Universal Robots URScript: FeedConveyor.script

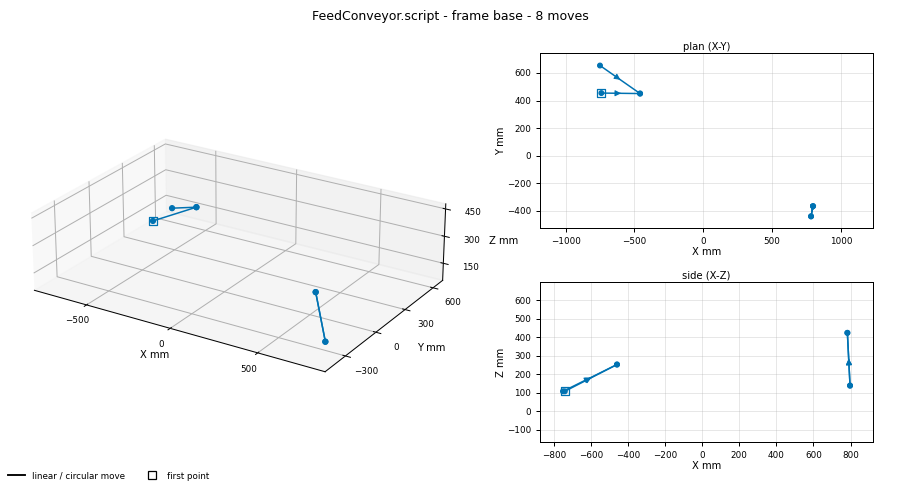
[picture p0: tool path of FeedConveyor.script in frame base, 8 of 12 moves have a stored position in this frame; points joined in program order, loops and branches not executed]
def FeedConveyor():
  # Global parameters:
  global speed_ms    = 0.250
  global speed_rads  = 0.750
  global accel_mss   = 1.200
  global accel_radss = 1.200
  global blend_radius_m = 0.001
  global ref_frame = p[0,0,0,0,0,0]

  #
  # TO REMOVE HEADER:
  # Go to "Program" -> "Post-Processor Editor"
  # Select "Universal Robots"
  # Set "INCLUDE_HEADER" to "False"
  #
  #--------------------------
  # Add any default subprograms here
  # For example, to drive a gripper as a program call:
  # def Gripper_Open():
  #   ...
  # end
  #
  # Example to drive a spray gun:
  def SprayOn(value):
    # use the value as an output:
    DO_SPRAY = 5
    if value == 0:
      set_standard_digital_out(DO_SPRAY, False)
    else:
      set_standard_digital_out(DO_SPRAY, True)
    end
  end

  # Example to drive an extruder:
  def Extruder(value):
    # use the value as an output:
    if value < 0:
      # stop extruder
    else:
      # start extruder
    end
  end

  # Example to move an external axis
  def MoveAxis(value):
    # use the value as an output:
    DO_AXIS_1 = 1
    DI_AXIS_1 = 1
    if value <= 0:
      set_standard_digital_out(DO_AXIS_1, False)

      # Wait for digital input to change state
      #while (get_standard_digital_in(DI_AXIS_1) != False):
      #  sync()
      #end
    else:
      set_standard_digital_out(DO_AXIS_1, True)

      # Wait for digital input to change state
      #while (get_standard_digital_in(DI_AXIS_1) != True):
      #  sync()
      #end
    end
  end
  #--------------------------


  # Main program:
  # Program generated by VerticalBot Studio for UR10 A on 25/10/2026 12:00:00
  # Using nominal kinematics.
  ref_frame = p[-1.052120, 0.561703, 0.068352, 0.000000, 0.000000, 1.570796]
  set_tcp(p[0.000000, -0.020000, 0.130000, 0.000000, 0.000000, 0.000000])
  movej([-1.414502, -1.531893, 2.172743, -0.640850, 0.156295, 0.000000],accel_radss,speed_rads,0,0.001)
  movel(pose_trans(ref_frame,p[-0.107464, -0.311695, 0.040000, 0.000000, 2.221441, 2.221441]),accel_mss,speed_ms,0,0.001)
  # Attach to GripperA Opened
  sleep(0.500)
  movel(pose_trans(ref_frame,p[-0.111072, -0.592992, 0.184438, -0.000000, -2.221441, -2.221441]),accel_mss,speed_ms,0,0.001)
  movej([2.282489, -0.754382, 0.716212, 0.038171, -0.885442, -0.000000],accel_radss,speed_rads,0,0.001)
  ref_frame = p[0.597228, -0.467251, 0.119180, 0.000000, 0.000000, 0.000000]
  movel(pose_trans(ref_frame,p[0.200000, 0.100000, 0.020000, -0.000000, 2.221441, 2.221441]),accel_mss,speed_ms,0,0.001)
  # Detach from GripperA Opened
  sleep(0.500)
  movel(pose_trans(ref_frame,p[0.185681, 0.025792, 0.304534, 0.029080, -2.208177, -2.208177]),accel_mss,speed_ms,0,0.001)
  movej([-1.414502, -1.531893, 2.172743, -0.640850, 0.156295, 0.000000],accel_radss,speed_rads,0,0.001)
  ref_frame = p[-1.052120, 0.561703, 0.068352, 0.000000, 0.000000, 1.570796]
  movel(pose_trans(ref_frame,p[0.092552, -0.301726, 0.040000, 0.000000, 2.221441, 2.221441]),accel_mss,speed_ms,0,0.001)
  # Attach to GripperA Opened
  sleep(0.500)
  movel(pose_trans(ref_frame,p[-0.111072, -0.592992, 0.184438, -0.000000, -2.221441, -2.221441]),accel_mss,speed_ms,0,0.001)
  movej([2.282489, -0.754382, 0.716212, 0.038171, -0.885442, -0.000000],accel_radss,speed_rads,0,0.001)
  ref_frame = p[0.597228, -0.467251, 0.119180, 0.000000, 0.000000, 0.000000]
  movel(pose_trans(ref_frame,p[0.200000, 0.100000, 0.020000, -0.000000, 2.221441, 2.221441]),accel_mss,speed_ms,0,0.001)
  # Detach from GripperA Opened
  sleep(0.500)
  movel(pose_trans(ref_frame,p[0.185681, 0.025792, 0.304534, 0.029080, -2.208177, -2.208177]),accel_mss,speed_ms,0,0.001)
  # End of main program
end

FeedConveyor()
